Staubli VAL3: copy.pgx

public program copy(string x_sKey, bool& x_bToSave)
  local bool l_bResult
  local string l_sName
begin
  if x_sKey!=""
    l_bResult=userPagePrompt("复制-输入新名称：",l_sName)
    if l_bResult
      if !isDefined(progTemp:pProgItem[l_sName])
        insert(progTemp:pProgItem[l_sName])
        call copyItem(l_sName,x_sKey)

        x_bToSave=true
      else
        userPageAlert("存在相同名称的程序！")
      endIf
    endIf
  endIf
end
